(* IEC 61131-3 sources: codesys-to-astra/tools/tests/fixtures/sourcemap/src/POUs/FB_Probe, 5 files *)

(* ---- FB_Probe.decl.st ---- *)
FUNCTION_BLOCK FB_Probe IMPLEMENTS I_Prio
VAR
    afbT : ARRAY[0..GVL_Const.SLOTS_MAX - 1] OF TON;
    aaiGrid : ARRAY[0..1] OF
        ARRAY[0..2] OF INT;
    astP : ARRAY[0..1] OF ST_Probe;   // @6
    iSlot : INT := 0;                 // @7
    rX : REAL := 0.0;
    xQ : BOOL := FALSE;
    tT : TIME := T#0S;
    iPrio : INT := 0;
    wMask : WORD := WORD#16#FF;       // @12
END_VAR

(* ---- FB_Probe.impl.st ---- *)
IF rX = 1.5 THEN rX := 0.0; ELSE rX := 1.0; END_IF   // @1
aaiGrid[iSlot,
        0] := 1;
IF rX = 1.5 THEN rX := 0.0; ELSE rX := 1.0; END_IF   // @4
xQ := afbT[iSlot]
    .Q;
IF rX = 1.5 THEN rX := 0.0; ELSE rX := 1.0; END_IF   // @7
afbT[iSlot](IN := TRUE,
            PT := T#1h500ms);
IF rX = 1.5 THEN rX := 0.0; ELSE rX := 1.0; END_IF   // @10
rX := astP[iSlot]
    .rLim;
IF rX = 1.5 THEN rX := 0.0; ELSE rX := 1.0; END_IF   // @13
IF xQ THEN
    ;
ELSE
END_IF
IF rX = 1.5 THEN rX := 0.0; ELSE rX := 1.0; END_IF   // @18
tT := TIME(
);
IF rX = 1.5 THEN rX := 0.0; ELSE rX := 1.0; END_IF   // @21
CASE iSlot OF
    0:
    1: xQ := TRUE;;
ELSE
END_CASE
IF rX = 1.5 THEN rX := 0.0; ELSE rX := 1.0; END_IF   // @27
xQ := xQ AND_THEN
    (rX > 0.0);
IF rX = 1.5 THEN rX := 0.0; ELSE rX := 1.0; END_IF   // @30
aaiGrid[0]
    [iSlot] := 2;
IF rX = 1.5 THEN rX := 0.0; ELSE rX := 1.0; END_IF   // @33
afbT[iSlot
    ](IN := FALSE);
if rX = 1.5 then rX := 0.0; else rX := 1.0; end_if   // @36
IF tT = TIME() THEN xQ := TRUE; ELSE xQ := FALSE; END_IF   // @37

(* ---- Priority.get.impl.st ---- *)
Priority := iPrio;
IF rX = 1.5 THEN rX := 0.0; ELSE rX := 1.0; END_IF   // @2

(* ---- Run.method.decl.st ---- *)
METHOD Run : BOOL
VAR_INPUT
    aiIn : ARRAY[0..GVL_Const.SLOTS_MAX
        - 1] OF INT;
END_VAR
VAR
    rY : REAL := 0.0;   // @7
END_VAR

(* ---- Run.method.impl.st ---- *)
IF rY = 1.5 THEN rY := 0.0; ELSE rY := 1.0; END_IF   // @1
rY := astP[iSlot].arStep[1]
    + astP[0].rLim;
IF rY = 1.5 THEN rY := 0.0; ELSE rY := 1.0; END_IF   // @4
WHILE FALSE DO
END_WHILE
IF rY = 1.5 THEN rY := 0.0; ELSE rY := 1.0; END_IF   // @7
Run := TRUE;
